LAYER Default
  FBS
    ProcessingStat : Processing2CAT;
    ProcHandling : TransportHandlingCAT;
    Station2 : Waypoint(skipStation := FALSE);
    Station1 : Waypoint(skipStation := FALSE);
    Station3 : Waypoint(skipStation := TRUE);
    Station4 : Waypoint(skipStation := FALSE);
    Station5 : Waypoint(skipStation := TRUE);
    Station6 : Waypoint(skipStation := FALSE);
    Distribution : Distribution2CAT;
    FB1 : TestingStation;
    TG1 : TransportGeneral1;
    OutputSorting : Sorting;
    OutputHanding : OutputHanding;
    RobotsStation : RoboCat;
    SB0 : LampControl(address := http://10.135.109.113/do_value/slot_0);
    CapDist : CapDistributionCAT;
  END_FBS
  EVENT_CONNECTIONS
    TG1.D8843CC7A5B75494 TO SB0.392A47A15328CAF8;
    ProcHandling.188659C343A79824 TO SB0.8038AD690A2EBB6D;
    ProcHandling.8A009C673F50EDC2 TO SB0.65194209493D291A;
    FB1.84F904613E536B04 TO SB0.7AA27EB4D48AA0EF;
    FB1.2A10A5926A92C41B TO SB0.37D71EDEC4A1963A;
    OutputHanding.B5C8731F109F88CC TO SB0.FAC1B651F864C1B0;
    OutputHanding.D930A57251D24EB8 TO SB0.7D58E289E5580604;
    RobotsStation.A39BFC97654CAFF3 TO CapDist.E4C6FDAF265EC198;
  END_CONNECTIONS
  ADAPTER_CONNECTIONS
    ProcessingStat.51D700913D16FC9C TO ProcHandling.43CECDD8B0A4C762;
    Distribution.1FE7610F8BFD7357 TO FB1.37BEEDB51F13C1BE;
    FB1.E98DD27C7D9BB7CB TO Station1.95F185C12A487DCF;
    ProcHandling.FFB46226821095B6 TO Station2.95F185C12A487DCF;
    Station3.54FF2A728F5BD4E9 TO TG1.64BF5537CA04CC7F;
    Station2.54FF2A728F5BD4E9 TO TG1.D21C0433245314C3;
    Station1.54FF2A728F5BD4E9 TO TG1.898CCF337DAF8974;
    Station6.54FF2A728F5BD4E9 TO TG1.C30F5862E83BFD5F;
    Station5.54FF2A728F5BD4E9 TO TG1.DC4A9CA3278BB557;
    Station4.54FF2A728F5BD4E9 TO TG1.4D4FE9F8A61F9CEC;
    OutputSorting.628B8F7074D40D3F TO OutputHanding.0A5D8ECE28FE65D8;
    OutputHanding.08D8FD6E7A0C852A TO Station6.95F185C12A487DCF;
    RobotsStation.1ED8A73DA6B21594 TO Station4.95F185C12A487DCF;
  END_CONNECTIONS
END_LAYER
